(* PLC project  *)
(* stored: creationDateTime 2026-04-10T12:42:14.376, modificationDateTime 2026-04-10T12:42:14.376 *)

{attribute 'qualified_only'}
{attribute 'strict'}
TYPE bds_snsrPr4_inst_te : (pSnsr_E := 0, bds_snsrPr4_numInst_E) USINT;
END_TYPE

{attribute 'qualified_only'}
{attribute 'strict'}
TYPE bds_snsrDst_inst_te : (SpdSnsr_E := 0, bds_snsrDst_numInst_E) USINT;
END_TYPE

{attribute 'qualified_only'}
{attribute 'strict'}
TYPE bds_snsrDsa_inst_te : (bds_snsrDsa_numInst_E) USINT;
END_TYPE

{attribute 'qualified_only'}
{attribute 'strict'}
TYPE bds_snsrPal_inst_te : (bds_snsrPal_numInst_E) USINT;
END_TYPE

{attribute 'qualified_only'}
{attribute 'strict'}
TYPE bds_in_aiv_signal_te : (IN_AIV_START_SIGNALS := 16#500, IN_AIV_START := 16#4FF, K52, K60, K43, K54, K55, K39, K38, K40, K42, K37, K61, K45, K44, A21, A36, A37, A38, A39, K30, A43, A22, A23, A24, K78, K76, K74, K77, K10, K75, K31, K34, A13, A40, A41, A42, A25, A26, A27, A14, A57, A28, A29, K11, K35, IN_AIV_NUM_SIGNALS, IN_AIV_FLEXIN_NUM_SIGNALS := K78) UINT;
END_TYPE

{attribute 'qualified_only'}
{attribute 'strict'}
TYPE bds_out_aov_signal_te : (OUT_AOV_START_SIGNALS := 16#300, OUT_AOV_START := 16#2FF, K25, A12, K62, OUT_AOV_NUM_SIGNALS, OUT_AOV_PVG_NUM_SIGNALS := K62) UINT;
END_TYPE

{attribute 'qualified_only'}
{attribute 'strict'}
TYPE bds_outClcU_signal_te : (bds_outClcU_K25_E := 0, bds_outClcU_A12_E, bds_outClcU_K62_E, bds_outClcU_numSignal_E) USINT;
END_TYPE

{attribute 'qualified_only'}
{attribute 'strict'}
TYPE bds_sys_ait_signal_te : (SYS_AIT_START_SIGNALS := 16#900, SYS_AIT_START := 16#8FF, TSGI1, TSGI2, SYS_AIT_NUM_SIGNALS) UINT;
END_TYPE

{attribute 'qualified_only'}
{attribute 'strict'}
TYPE bds_in_di_signal_te : (IN_DI_START_SIGNALS := 16#400, IN_DI_START := 16#3FF, K22, K21, IN_DI_NUM_SIGNALS) UINT;
END_TYPE

{attribute 'qualified_only'}
{attribute 'strict'}
TYPE bds_in_ri_signal_te : (IN_RI_START_SIGNALS := 16#600, IN_RI_START := 16#5FF, K41, K65, K63, K64, K32, K33, IN_RI_NUM_SIGNALS) UINT;
END_TYPE

{attribute 'qualified_only'}
{attribute 'strict'}
TYPE bds_in_fi_signal_te : (IN_FI_START_SIGNALS := 16#700, IN_FI_START := 16#6FF, K39_VI, K38_VI, K40_VI, K41_VI, K42_VI, K45_VI, K44_VI, K65_VI, K63_VI, K64_VI, A36_VI, A37_VI, A38_VI, A39_VI, K54_VI, K37_VI, K30_VI, A43_VI, IN_FI_NUM_SIGNALS, IN_FI_DSM_NUM_SIGNALS := IN_FI_NUM_SIGNALS) UINT;
END_TYPE

{attribute 'qualified_only'}
{attribute 'strict'}
TYPE bds_in_sent_signal_te : (IN_SENT_START_SIGNALS := 16#800, IN_SENT_START := 16#7FF, K53, K59, K57, K58, K36, K56, IN_SENT_NUM_SIGNALS) UINT;
END_TYPE

{attribute 'qualified_only'}
{attribute 'strict'}
TYPE bds_in_phase_signal_te : (IN_PHASE_START_SIGNALS := 16#900, IN_PHASE_START := 16#8FF, K55_VI_K61_VI, IN_PHASE_NUM_SIGNALS) UINT;
END_TYPE

{attribute 'qualified_only'}
{attribute 'strict'}
TYPE bds_out_do_signal_te : (OUT_DO_START_SIGNALS := 16#100, OUT_DO_START := 16#FF, K13, A04, A10, A56, A11, A55, A01, A06, A16, A58, A49, A50, K84, K85, K86, K87, OUT_DO_NUM_SIGNALS, OUT_DO_FSC_NUM_SIGNALS := K84) UINT;
END_TYPE

{attribute 'qualified_only'}
{attribute 'strict'}
TYPE bds_out_po_signal_te : (OUT_PO_START_SIGNALS := 16#200, OUT_PO_START := 16#1FF, K07, K09, K73, K08, K29, K17, A32, A47, A31, A48, A46, A33, A34, A51, A35, A53, A52, A54, K16, K14, K15, A19, A05, A20, A09, A02, A17, K51, K12, A03, A18, A08, A07, K80, K81, K82, K83, OUT_PO_NUM_SIGNALS, OUT_PO_FSC_NUM_SIGNALS := K80, OUT_PO_FSC_HS_NUM_SIGNALS := K16) UINT;
END_TYPE

{attribute 'external_name' := 'cmp_rts_bds_outDig_signal_te'}
TYPE bds_outDig_signal_te : (bds_outDig_K13_E := 0, bds_outDig_A04_E, bds_outDig_A10_E, bds_outDig_A56_E, bds_outDig_A11_E, bds_outDig_A55_E, bds_outDig_A01_E, bds_outDig_A06_E, bds_outDig_A16_E, bds_outDig_A58_E, bds_outDig_A49_E, bds_outDig_A50_E, bds_outDig_K84_E, bds_outDig_K85_E, bds_outDig_K86_E, bds_outDig_K87_E, bds_outDig_K07_E, bds_outDig_K09_E, bds_outDig_K73_E, bds_outDig_K08_E, bds_outDig_K29_E, bds_outDig_K17_E, bds_outDig_A32_E, bds_outDig_A47_E, bds_outDig_A31_E, bds_outDig_A48_E, bds_outDig_A46_E, bds_outDig_A33_E, bds_outDig_A34_E, bds_outDig_A51_E, bds_outDig_A35_E, bds_outDig_A53_E, bds_outDig_A52_E, bds_outDig_A54_E, bds_outDig_K16_E, bds_outDig_K14_E, bds_outDig_K15_E, bds_outDig_A19_E, bds_outDig_A05_E, bds_outDig_A20_E, bds_outDig_A09_E, bds_outDig_A02_E, bds_outDig_A17_E, bds_outDig_K51_E, bds_outDig_K12_E, bds_outDig_A03_E, bds_outDig_A18_E, bds_outDig_A08_E, bds_outDig_A07_E, bds_outDig_K80_E, bds_outDig_K81_E, bds_outDig_K82_E, bds_outDig_K83_E, bds_outDig_numSignal_E) USINT;
END_TYPE

{attribute 'external_name' := 'cmp_rts_bds_outPwm_signal_te'}
TYPE bds_outPwm_signal_te : (bds_outPwm_K07_E := 0, bds_outPwm_K09_E, bds_outPwm_K73_E, bds_outPwm_K08_E, bds_outPwm_K29_E, bds_outPwm_K17_E, bds_outPwm_A32_E, bds_outPwm_A47_E, bds_outPwm_A31_E, bds_outPwm_A48_E, bds_outPwm_A46_E, bds_outPwm_A33_E, bds_outPwm_A34_E, bds_outPwm_A51_E, bds_outPwm_A35_E, bds_outPwm_A53_E, bds_outPwm_A52_E, bds_outPwm_A54_E, bds_outPwm_K16_E, bds_outPwm_K14_E, bds_outPwm_K15_E, bds_outPwm_A19_E, bds_outPwm_A05_E, bds_outPwm_A20_E, bds_outPwm_A09_E, bds_outPwm_A02_E, bds_outPwm_A17_E, bds_outPwm_K51_E, bds_outPwm_K12_E, bds_outPwm_A03_E, bds_outPwm_A18_E, bds_outPwm_A08_E, bds_outPwm_A07_E, bds_outPwm_K80_E, bds_outPwm_K81_E, bds_outPwm_K82_E, bds_outPwm_K83_E, bds_outPwm_numSignal_E) USINT;
END_TYPE

{attribute 'qualified_only'}
{attribute 'strict'}
TYPE bds_sys_aiv_signal_te : (SYS_AIV_START_SIGNALS := 16#A00, SYS_AIV_START := 16#9FF, UBAT_MON, UBRM24_MON, VDD5A_MON, UBR24_VP, UBRM24_LOADS, VDD3V3, VPR6, VDD5V_IN, VDD5_S3530, VSS3V5, VSS4V10, LSS_MEAS_CL13, LSS_MEAS_CL2, SYS_AIV_NUM_SIGNALS) UINT;
END_TYPE

{attribute 'qualified_only'}
{attribute 'strict'}
TYPE bds_sys_do_signal_te : (SYS_DO_START_SIGNALS := 16#B00, SYS_DO_START := 16#AFF, SHUNT_AIC_K39_EN, SHUNT_AIC_K38_EN, SHUNT_AIC_K40_EN, SHUNT_AIC_K41_EN, SHUNT_AIC_K42_EN, SHUNT_AIC_K45_EN, SHUNT_AIC_K44_EN, SHUNT_AIC_K65_EN, SHUNT_AIC_K63_EN, SHUNT_AIC_K64_EN, SHUNT_AIC_A36_EN, SHUNT_AIC_A37_EN, SHUNT_AIC_A38_EN, SHUNT_AIC_A39_EN, SHUNT1_EN, SHUNT3_EN, SHUNT5_EN, SHUNT6_EN, SYS_DO_NUM_SIGNALS) UINT;
END_TYPE

{attribute 'qualified_only'}
{attribute 'strict'}
TYPE bds_sys_vss_signal_te : (SYS_VSS_START_SIGNALS := 16#C00, SYS_VSS_START := 16#BFF, VSS1, VSS2, VSS3, VSS4, SYS_VSS_NUM_SIGNALS, SYS_VSS_CY_NUM_SIGNALS := VSS3) UINT;
END_TYPE

{attribute 'qualified_only'}
{attribute 'strict'}
TYPE bds_sys_di_signal_te : (SYS_DI_START_SIGNALS := 16#D00, SYS_DI_START := 16#CFF, ST_INH, SYS_DI_NUM_SIGNALS) UINT;
END_TYPE

{attribute 'qualified_only'}
{attribute 'strict'}
TYPE bds_snsrPr4_inst_te : (pSnsr_E := 0, bds_snsrPr4_numInst_E) USINT;
END_TYPE

{attribute 'qualified_only'}
{attribute 'strict'}
TYPE bds_snsrDst_inst_te : (SpdSnsr_E := 0, bds_snsrDst_numInst_E) USINT;
END_TYPE

{attribute 'qualified_only'}
{attribute 'strict'}
TYPE bds_snsrDsa_inst_te : (bds_snsrDsa_numInst_E := 0) USINT;
END_TYPE

{attribute 'qualified_only'}
{attribute 'strict'}
TYPE bds_snsrPal_inst_te : (bds_snsrPal_numInst_E := 0) USINT;
END_TYPE

(* Definition of input Configured Signals for Voltage( Consists signals of all variants) *)
{attribute 'qualified_only'}
{attribute 'strict'}
TYPE bds_inU_signal_te : (bds_inU_K52_E := 0, bds_inU_K60_E, bds_inU_K43_E, bds_inU_K54_E, bds_inU_K55_E, bds_inU_K39_E, bds_inU_K38_E, bds_inU_K40_E, bds_inU_K42_E, bds_inU_K37_E, bds_inU_K61_E, bds_inU_K45_E, bds_inU_K44_E, bds_inU_A21_E, bds_inU_A36_E, bds_inU_A37_E, bds_inU_A38_E, bds_inU_A39_E, bds_inU_K30_E, bds_inU_A43_E, bds_inU_A22_E, bds_inU_A23_E, bds_inU_A24_E, bds_inU_K78_E, bds_inU_K76_E, bds_inU_K74_E, bds_inU_K77_E, bds_inU_K10_E, bds_inU_K75_E, bds_inU_K31_E, bds_inU_K34_E, bds_inU_A13_E, bds_inU_A40_E, bds_inU_A41_E, bds_inU_A42_E, bds_inU_A25_E, bds_inU_A26_E, bds_inU_A27_E, bds_inU_A14_E, bds_inU_A57_E, bds_inU_A28_E, bds_inU_A29_E, bds_inU_K11_E, bds_inU_K35_E, bds_inU_A59_E, bds_inU_numSignal_E) USINT;
END_TYPE

(* values of bds_inDig_signal_te: bds_inDig_K21_E: End V1 *)

(* BODAS configuration of available digital input signals *)
{attribute 'qualified_only'}
{attribute 'strict'}
TYPE bds_inDig_signal_te : (bds_inDig_K22_E := 0, bds_inDig_K21_E, bds_inDig_numSignal_E) USINT;
END_TYPE

(* Definition of input signals for Resistance *)
{attribute 'qualified_only'}
{attribute 'strict'}
TYPE bds_inR_signal_te : (bds_inR_K41_E := 0, bds_inR_K65_E, bds_inR_K63_E, bds_inR_K64_E, bds_inR_K32_E, bds_inR_K33_E, bds_inR_numSignal_E) USINT;
END_TYPE

(* values of bds_sent_signal_te: bds_sent_K53_E: X_X_X03; bds_sent_K59_E: X_X_X04; bds_sent_K57_E: X_X_X16; bds_sent_K58_E: X_X_X17; bds_sent_K36_E: X_X_X18; bds_sent_K56_E: X_X_X19 *)

(* Definition configuration of available SENT signals (consists signals of all variants) *)
{attribute 'qualified_only'}
{attribute 'strict'}
TYPE bds_sent_signal_te : (bds_sent_K53_E := 0, bds_sent_K59_E, bds_sent_K57_E, bds_sent_K58_E, bds_sent_K36_E, bds_sent_K56_E, bds_sent_numSignal_E) USINT;
END_TYPE

(* Definition of input signals for PWM *)
{attribute 'qualified_only'}
{attribute 'strict'}
TYPE bds_inPwm_signal_te : (bds_inPwm_K54_E := 0, bds_inPwm_K37_E, bds_inPwm_K30_E, bds_inPwm_A43_E, bds_inPwm_A59_A44_E, bds_inPwm_numSignal_E) USINT;
END_TYPE

{attribute 'external_name' := 'cmp_rts_bds_inPha_signal_te'}
TYPE bds_inPha_signal_te : (bds_inPha_K55_K61_E := 0, bds_inPha_numSignal_E) USINT;
END_TYPE

(* values of bds_inI_signal_te: bds_inI_A43_E: End V1 *)

(* BODAS configuration of available current measurement input signals *)
{attribute 'qualified_only'}
{attribute 'strict'}
TYPE bds_inI_signal_te : (bds_inI_A38_E := 0, bds_inI_A39_E, bds_inI_K37_E, bds_inI_K30_E, bds_inI_A43_E, bds_inI_numSignal_E) USINT;
END_TYPE

(* post build system variants information *)
{attribute 'qualified_only'}
{attribute 'strict'}
TYPE bds_sysPb_vrnt_te : (bds_sysPb_vrnt01_E  := 0, bds_sysPb_maxNumVrnt_E) USINT;
END_TYPE

{attribute 'qualified_only'}
VAR_GLOBAL CONSTANT  (* bds_sysIo_ec_gvl *)
  BDS_SYSIO_FI_SHUNT_NUM_SIGNALS_D : UINT := bds_sys_do_signal_te.SHUNT1_EN;
END_VAR

{attribute 'qualified_only'}
VAR_GLOBAL CONSTANT  (* bds_in_legacy_ec_gvl *)
  ACTIVATE_SHUNT_AIC_K39 : UDINT := 0;
  ACTIVATE_SHUNT_AIC_K38 : UDINT := 0;
  ACTIVATE_SHUNT_AIC_K40 : UDINT := 0;
  ACTIVATE_SHUNT_AIC_K41 : UDINT := 0;
  ACTIVATE_SHUNT_AIC_K42 : UDINT := 0;
  ACTIVATE_SHUNT_AIC_K45 : UDINT := 0;
  ACTIVATE_SHUNT_AIC_K44 : UDINT := 0;
  ACTIVATE_SHUNT_AIC_K65 : UDINT := 0;
  ACTIVATE_SHUNT_AIC_K63 : UDINT := 0;
  ACTIVATE_SHUNT_AIC_K64 : UDINT := 0;
  ACTIVATE_SHUNT_AIC_A36 : UDINT := 0;
  ACTIVATE_SHUNT_AIC_A37 : UDINT := 0;
  ACTIVATE_SHUNT_AIC_A38 : UDINT := 1;
  ACTIVATE_SHUNT_AIC_A39 : UDINT := 1;
  ACTIVATE_SHUNT1 : UDINT := 0;
  ACTIVATE_SHUNT2 : UDINT := 0;
  ACTIVATE_SHUNT3 : UDINT := 1;
  ACTIVATE_SHUNT4 : UDINT := 0;
  ACTIVATE_SHUNT5 : UDINT := 1;
  ACTIVATE_SHUNT6 : UDINT := 1;
  BDS_IN_AIV_32V_NUM_SIGNALS_D : UINT := bds_in_aiv_signal_te.A14;
  BDS_IN_FI_AIC_NUM_SIGNALS_D : UINT := bds_in_fi_signal_te.K54_VI;
END_VAR

{attribute 'qualified_only'}
VAR_GLOBAL CONSTANT  (* bds_out_ec_gvl *)
  RECONF_X_X_X25 : UDINT := 0;
END_VAR

{attribute 'qualified_only'}
VAR_GLOBAL CONSTANT  (* bds_in_ec_gvl *)
  BDS_inCmn_postVariants_DU8 : USINT := 1;
END_VAR

{attribute 'qualified_only'}
VAR_GLOBAL CONSTANT  (* bds_sent_ec_gvl *)
  bds_sent_postVariants_du8 : USINT := 1;
  bds_sent_maxDataNibbles_du8 : USINT := 6;
  bds_sent_rxFastDataBufSize_du8 : USINT := 0;
  bds_sent_rxSlowDataBufSize_du8 : USINT := 0;
END_VAR

{attribute 'qualified_only'}
VAR_GLOBAL CONSTANT  (* bds_sysPb_ec_gvl *)
  ml290rts_bs_HelloWorld : USINT := bds_sysPb_vrnt_te.bds_sysPb_vrnt01_E;
END_VAR
